(* IEC 61131-3 sources: plcassist-cli/packages/volt-lsp-iec/test-corpus/awa-palletizer/Device/Plc Logic/Application/Library Manager/(unresolved)/l_st2i_activatetimemeasurement, 1 file *)

(* ---- GVL_TIMEMEASUREMENT.gvl ---- *)
VAR_GLOBAL
	XACTIVATETIMEMEASUREMENT : BOOL := FALSE;
END_VAR
